// Tests for FB_IagCabinet, the I_Cabinet with the physical Local/Remote key: key to control mode and the safety pass-through.
FUNCTION_BLOCK FB_IagCabinet_Tests EXTENDS TcUnit.FB_TestSuite
VAR
END_VAR

Key_Off_Is_Remote();
Key_On_Is_Local();
Mode_Follows_The_Key();
Switch_Is_Present();
Estop_Passes_Through();
Safety_Error_Passes_Through();
Ack_Pending_Passes_Through();
Pendant_Passes_Through_And_Is_Independent();

METHOD PRIVATE Key_Off_Is_Remote
VAR
	fbCabinet	: FB_IagCabinet;
END_VAR
TEST('Key_Off_Is_Remote');
fbCabinet(bLocalKey := FALSE);
AssertTrue(Condition := fbCabinet.ControlMode = E_ControlMode.remote, Message := 'remote');
TEST_FINISHED();
END_METHOD

METHOD PRIVATE Key_On_Is_Local
VAR
	fbCabinet	: FB_IagCabinet;
END_VAR
TEST('Key_On_Is_Local');
fbCabinet(bLocalKey := TRUE);
AssertTrue(Condition := fbCabinet.ControlMode = E_ControlMode.local, Message := 'local');
TEST_FINISHED();
END_METHOD

METHOD PRIVATE Mode_Follows_The_Key
VAR
	fbCabinet	: FB_IagCabinet;
END_VAR
TEST('Mode_Follows_The_Key');
fbCabinet(bLocalKey := TRUE);
fbCabinet(bLocalKey := FALSE);
AssertTrue(Condition := fbCabinet.ControlMode = E_ControlMode.remote, Message := 'back to remote');
TEST_FINISHED();
END_METHOD

METHOD PRIVATE Switch_Is_Present
VAR
	fbCabinet	: FB_IagCabinet;
END_VAR
TEST('Switch_Is_Present');
fbCabinet(bLocalKey := FALSE);
AssertTrue(Condition := fbCabinet.SwitchPresent, Message := 'switch present, key off');
fbCabinet(bLocalKey := TRUE);
AssertTrue(Condition := fbCabinet.SwitchPresent, Message := 'switch present, key on');
TEST_FINISHED();
END_METHOD

METHOD PRIVATE Estop_Passes_Through
VAR
	fbCabinet	: FB_IagCabinet;
END_VAR
TEST('Estop_Passes_Through');
fbCabinet(bEstop := FALSE);
AssertFalse(Condition := fbCabinet.EstopActive, Message := 'no e-stop');
fbCabinet(bEstop := TRUE);
AssertTrue(Condition := fbCabinet.EstopActive, Message := 'e-stop');
TEST_FINISHED();
END_METHOD

METHOD PRIVATE Safety_Error_Passes_Through
VAR
	fbCabinet	: FB_IagCabinet;
END_VAR
TEST('Safety_Error_Passes_Through');
fbCabinet(bSafetyError := FALSE);
AssertFalse(Condition := fbCabinet.SafetyError, Message := 'no error');
fbCabinet(bSafetyError := TRUE);
AssertTrue(Condition := fbCabinet.SafetyError, Message := 'error');
TEST_FINISHED();
END_METHOD

METHOD PRIVATE Ack_Pending_Passes_Through
VAR
	fbCabinet	: FB_IagCabinet;
END_VAR
TEST('Ack_Pending_Passes_Through');
fbCabinet(bSafetyAckPending := FALSE);
AssertFalse(Condition := fbCabinet.SafetyAckPending, Message := 'no ack pending');
fbCabinet(bSafetyAckPending := TRUE);
AssertTrue(Condition := fbCabinet.SafetyAckPending, Message := 'ack pending');
TEST_FINISHED();
END_METHOD

METHOD PRIVATE Pendant_Passes_Through_And_Is_Independent
VAR
	fbCabinet	: FB_IagCabinet;
END_VAR
TEST('Pendant_Passes_Through_And_Is_Independent');
fbCabinet(bLocalKey := TRUE, bPendantActive := FALSE);
AssertFalse(Condition := fbCabinet.PendantActive, Message := 'no pendant');
fbCabinet(bLocalKey := FALSE, bPendantActive := TRUE);
AssertTrue(Condition := fbCabinet.PendantActive, Message := 'pendant');
AssertFalse(Condition := fbCabinet.EstopActive, Message := 'other signals untouched');
TEST_FINISHED();
END_METHOD

END_FUNCTION_BLOCK

(* stored: Version 1.1.0.1, ProductVersion 3.1.4024.15
   POU FB_IagCabinet_Tests: Id {2c4fdf76-ff0e-413b-b54b-092c338eacf4}, SpecialFunc None
   Method Key_Off_Is_Remote: Id {b44a8da9-fbe0-4161-b67e-ffd9def771d9}
   Method Key_On_Is_Local: Id {3a67a2c6-2031-48a2-9405-ed8ee7756bc4}
   Method Mode_Follows_The_Key: Id {ba521a62-d79e-46bf-a8c4-158292f594b2}
   Method Switch_Is_Present: Id {7058100b-2cc8-4cb3-abe9-4e30739a616c}
   Method Estop_Passes_Through: Id {4356b4ad-ca03-4c7e-8d35-1b2874a9b2b1}
   Method Safety_Error_Passes_Through: Id {baad3948-2599-455b-a6b3-a0e5d8f7901f}
   Method Ack_Pending_Passes_Through: Id {e5b761fa-238d-4dcb-bb29-991c0f149908}
   Method Pendant_Passes_Through_And_Is_Independent: Id {edbe0fb8-afad-4407-bea4-05b56ab3e283} *)
